{attribute 'no_assign'}
FUNCTION_BLOCK FB_LN_WTURBINE_LD0_LLN0 EXTENDS FB_AcsiCommonLogicalNodeClass
VAR_INPUT
	NamPlt: FB_DO_WTURBINE_LD0_LLN0_NamPlt := (sClass:='LPL', bLinkResult:=THIS^.AddDataToContainer(ipData:=NamPlt));
	Beh: FB_DO_WTURBINE_LD0_LLN0_Beh := (sClass:='ENS', bLinkResult:=THIS^.AddDataToContainer(ipData:=Beh));
	Health: FB_DO_WTURBINE_LD0_LLN0_Health := (sClass:='ENS', bLinkResult:=THIS^.AddDataToContainer(ipData:=Health));
	Mod_: FB_DO_WTURBINE_LD0_LLN0_Mod := (sObjectName:='Mod', sClass:='ENC', bLinkResult:=THIS^.AddDataToContainer(ipData:=Mod_));
END_VAR
VAR
END_VAR

END_FUNCTION_BLOCK

(* stored: Version 1.1.0.1
   POU FB_LN_WTURBINE_LD0_LLN0: Id {35e2917c-60da-4c1b-af55-ccf7f9e680dc}, SpecialFunc None *)
